(*
SPDX-FileCopyrightText: c 2026 Oleksandr Tiutyk <trofimich@gmail.com>
SPDX-License-Identifier: MIT
License: https://opensource.org/license/mit
*)

(*!
<summary>Checks normal-open input values and transition detection.</summary>
<description>
Uses a live case-owned automation parent and fresh local device fixtures on every run.
The scenario reads and writes ordinary simulated storage within one task cycle.
</description>
*)

{attribute 'no_assign'}
{attribute 'no_explicit_call' := 'do not call this function block directly'}
FUNCTION_BLOCK DigitalInputNormallyOpenTest EXTENDS TOF_Testing.SingleCycleTest
VAR_STAT
	{attribute 'hide'}
	_ClassName : STRING := __POUNAME();
END_VAR
VAR
	//! <summary>Live parent borrowed by the method-local simulated device.</summary>
	_AutomationRoot : MockAutomationController(name := "DevicesIORoot");
END_VAR

(*!
<summary>Checks normal-open input values and transition detection.</summary>
*)
METHOD PROTECTED ExecuteTest
VAR
	input : TOF_Devices_IO.DigitalInput(name := "DI_NO", parent := _AutomationRoot);
	rawInput : BOOL;
END_VAR
input.Initialize();
input.BindToIO(rawValue := rawInput);

Assert.ThatBool(
	actual := input.BoundToIO,
	message := "DigitalInput should be bound to IO"
).IsTrue();

rawInput := FALSE;
input.ProcessInput();
Assert.ThatBool(
	actual := input.Value,
	message := "Value should be FALSE"
).IsFalse();

rawInput := TRUE;
input.ProcessInput();
Assert.ThatBool(
	actual := input.Value,
	message := "Value should be TRUE"
).IsTrue();
Assert.ThatBool(
	actual := input.Changed,
	message := "Changed should be TRUE on transition"
).IsTrue();

input.ProcessInput();
Assert.ThatBool(
	actual := input.Changed,
	message := "Changed should be FALSE when state remains same"
).IsFalse();
END_METHOD

//! <summary>Borrows the concrete class name. Callers must not modify it.</summary>
{attribute 'monitoring' := 'call'}
PROPERTY ClassName : REFERENCE TO STRING
GET
ClassName REF= _ClassName;
END_GET
END_PROPERTY

//! <summary>Borrows the compiler-initialized namespace name. Callers must not modify it.</summary>
{attribute 'monitoring' := 'call'}
PROPERTY NamespaceName : REFERENCE TO STRING
GET
NamespaceName REF= CurrentNamespace.Name;
END_GET
END_PROPERTY

//! <summary>Reports the concrete instance size in bytes.</summary>
{attribute 'monitoring' := 'call'}
PROPERTY SelfSize : ULINT
GET
SelfSize := XSIZEOF(THIS^);
END_GET
END_PROPERTY

END_FUNCTION_BLOCK

(* stored: Version 1.1.0.1
   POU DigitalInputNormallyOpenTest: Id {b47ab2fd-5062-493e-9b5b-24667747283e}, SpecialFunc None
   Method ExecuteTest: Id {a8b041d0-78f3-4389-adaa-8942723430d0}
   Property ClassName: Id {262355ac-351e-4112-aaad-b3eca7e9c55e}
   Get Get: Id {3b639424-2df2-4f0d-a9a5-63c02cb39136}
   Property NamespaceName: Id {a5157fc2-c3d5-405b-94db-3184b6e7fcf3}
   Get Get: Id {a6351aae-ed4d-44d4-a6e5-37bb1306ad35}
   Property SelfSize: Id {d3646eb8-c82f-4fb0-805f-19e885db6607}
   Get Get: Id {492eeb49-43f6-486f-99f4-74f3a71bc33e} *)
